Fanuc KAREL source: kt00739.KL

-- PROVISIONAL review KL for V770-1; original PC SHA256 b1e741a2de9c1c2321df2728878ad7b96a97476381bbe58dbdb5426220f39400
-- Incomplete behavior may be omitted. Consult companion uncertainty JSON. Do not deploy.
PROGRAM KT00739
%NOLOCKGROUP
VAR
  OUT : INTEGER
-- UNRESOLVED_DECL ARG type=002018
BEGIN
  -- UNRESOLVED_PC offsets 5-18; opcodes 22,1D,23
  -- UNRESOLVED_PC offsets 23-27; opcodes 7F
END KT00739
